Fanuc KAREL source: kb00128.KL

-- PROVISIONAL review KL for V770-1; original PC SHA256 e3e05ebc5381f77644f454d5b05750329ef269e2f25cd745647b1262c42f0adc
-- Incomplete behavior may be omitted. Consult companion uncertainty JSON. Do not deploy.
PROGRAM KB00128
%NOLOCKGROUP
BEGIN
  -- UNRESOLVED_PC offsets 5-28; opcodes 27,22,1C,31,4A
  -- UNRESOLVED_PC offsets 33-37; opcodes 7F
END KB00128
